// TIA Portal V19 export
DATA_BLOCK "ALL_AI_DB_1"   // DB16
// stored: InstanceOfName ALL_AI, InstanceOfType FB
"ALL_AI"
   // VAR
   //    AI_TT01 { S7_SetPoint := 'True'} : "AI";
   //    TT_01 { S7_SetPoint := 'True'} : "AI";
   //    TT_02 { S7_SetPoint := 'True'} : "AI";
   //    TT_03 { S7_SetPoint := 'True'} : "AI";
   //    APT01 { S7_SetPoint := 'True'} : "AI";
   //    GPT01 { S7_SetPoint := 'True'} : "AI";
   //    GPT02 { S7_SetPoint := 'True'} : "AI";
   //    GPT03 { S7_SetPoint := 'True'} : "AI";
   //    GPT04 { S7_SetPoint := 'True'} : "AI";
   //    O201 { S7_SetPoint := 'True'} : "AI";
   //    LEL01 { S7_SetPoint := 'True'} : "AI";
   //    LEL02 { S7_SetPoint := 'True'} : "AI";
   //    PS01 { S7_SetPoint := 'True'} : "AI";
   //    RLT01 { S7_SetPoint := 'True'} : "AI";
   //    Weighing { S7_SetPoint := 'True'} : "AI";
   // END_VAR
BEGIN
END_DATA_BLOCK
